(* IEC 61131-3 sources: SortJet_MasterSPS_Aufbau.fbsproj/09_Station/Stationen/_Basic/Basic_Schnittstelle_FB_V01_00_00.fb.st^, 6 files *)

(* ---- A_Changelog.act.st ---- *)
(* METADATA
{
	"v3Meta": {
		"objectGuid": "30bc6851-70b4-468b-8947-0ecaf15505c8"
	}
}
*)
{attribute 'excludefrombuild'}
ACTION A_Changelog
(* !!! VERSIONSÄNDERUNGEN WERDEN HIER DETAILLIERT DOKUMENTIERT !!!

- 2026-11-24 - V01_00_00: Tobias Brekerbohm
  - Erste Freigabe SortJet-Master
*)
END_ACTION

(* ---- A_Schnittstelle.act.st ---- *)
(* METADATA
{
	"v3Meta": {
		"objectGuid": "8ef5bc36-5f76-46e1-a5ac-606d922f719c"
	}
}
*)
ACTION A_Schnittstelle
//-------------------------------------------------------------------------------------------------
// AKTION SCHNITTSTELLE
//-------------------------------------------------------------------------------------------------

BasisStationsParameter.OutGlasTransport[cWAND_1].stStationsNummern          := BasisStationsParameter.stMKs.stStationsNummern;
BasisStationsParameter.OutGlasTransport[cWAND_1].wStationsTyp               := BasisStationsParameter.stMKs.eStationsTyp;
BasisStationsParameter.OutGlasTransport[cWAND_1].rLaengeStation             := BasisStationsParameter.stMKs.stFremdanlage.rLaengeStation;
BasisStationsParameter.OutGlasTransport[cWAND_1].bEinlaufsensor             REF= bEmpfaengerSensorEinlauf;
BasisStationsParameter.OutGlasTransport[cWAND_1].bAuslaufsensor             REF= bgFALSE;
BasisStationsParameter.OutGlasTransport[cWAND_1].bBereitZumAustransport     REF= blBereitZumAustransport;
BasisStationsParameter.OutGlasTransport[cWAND_1].bBereitZumEintransport     REF= blBereitZumEintransport;
BasisStationsParameter.OutGlasTransport[cWAND_1].rGeschwindigkeit           REF= rpGeschwindigkeit;
BasisStationsParameter.OutGlasTransport[cWAND_1].bFehler                    REF= BasisStationsParameter.bFehler;
BasisStationsParameter.OutGlasTransport[cWAND_1].bQuittScheibe              REF= bgFALSE;
BasisStationsParameter.OutGlasTransport[cWAND_1].bFreigabe                  REF= BasisStationsParameter.stFreigabe.bAlles;
BasisStationsParameter.OutGlasTransport[cWAND_1].bTransportAbgeschlossen    REF= bgFALSE;
BasisStationsParameter.OutGlasTransport[cWAND_1].bScheibeFaehrtUeberEinlauf REF= bgFALSE;
BasisStationsParameter.OutGlasTransport[cWAND_1].bScheibeFaehrtUeberAuslauf REF= bgFALSE;
BasisStationsParameter.OutGlasTransport[cWAND_1].bAutomatikBetriebAktiv     REF= blAutomatikBetriebAktiv;

//   - Status der Sortierung [Hardware- Ausgaenge]
//     => Automatik ativ
//     => Kein Fehler aktiv
out_bSenderBereit := blSenderBereit :=         BasisStationsParameter.bAutomatik
                     AND NOT BasisStationsParameter.bFehler
                     AND NOT BasisStationsParameter.InGlasTransportVorgaenger[cWAND_1].bFehler;

out_bSenderGlasBereit := blSenderGlasBereit (*OR bgVisu_Schnittstelle_GlasBereit[BasisStationsParameter.stMKs.stStationsNummern.NummerSPS]*);

// Eingangssignale können über den Drive oder IO's kommen
bEmpfaengerSensorEinlauf := bpEmpfaengerSensorEinlauf OR in_bEmpfaengerSensorEinlauf;

//-------------------------------------------------------------------------------------------------
// VISU
//-------------------------------------------------------------------------------------------------
bgVisu_Schnittstelle_GlasBereit[BasisStationsParameter.stMKs.stStationsNummern.NummerSPS]    := out_bSenderGlasBereit;
END_ACTION

(* ---- IGLineEvent.act.st ---- *)
(* METADATA
{
	"v3Meta": {
		"objectGuid": "eb410a9f-4f2d-4b91-9b42-1e80fc6ee1dd"
	}
}
*)
ACTION IGLineEvent
//-------------------------------------------------------------------------------------------------
// IG LINE EVENT
//-------------------------------------------------------------------------------------------------
bpISOLineEventAktiv := blUebergabeGlas;
(* Hinweis:
   - Ausgaenge setzen
*)
out_bLeuchteGlasbruch :=( blUebergabeGlas AND ((wpAuftragsTyp = 1) OR (wpAuftragsTyp = 4) OR ((wpAuftragsTyp = 5) AND gbFlashbit05sec))) ;
out_bLeuchteSpezial   :=( blUebergabeGlas AND ((wpAuftragsTyp = 2) OR ((wpAuftragsTyp = 3) AND gbFlashbit02sec )));

out_bAmpelEventAktiv := (blUebergabeGlas);

//-------------------------------------------------------------------------------------------------
// STEUERUNG:  ISO Line EVENT abhandeln
//-------------------------------------------------------------------------------------------------
IF ( bpStarteIGEvent
     AND NOT blUebergabeGlas )
THEN
  blUebergabeGlas := TRUE;
  bpStarteIGEvent := FALSE;
  steplUebergabeGlas := STEP_0_E;
END_IF

(* Hinweis:
   - wpAuftragsTyp:
   - case 0: //Kein Ereignis
   - case 1: //Scheibe von Isolinie abnehmen!
   - case 2: //Einschleusen von Sonderscheibe!
   - case 3: //Laufende!
   - case 4: //Alle Scheiben der Isoeinheit sind Bruch!
   - case 5: //Eine Scheibe der Einheit ist Bruch!
*)
IF ( blUebergabeGlas ) THEN
  CASE steplUebergabeGlas OF
    // GLASUEBERGABE ========================
    STEP_0_E:

      dwpWartezeit := 0;

      tlWarteZeiteAufnahme := TIME(); // Starten der Wartezeitenermittlung

      CASE wpAuftragsTyp OF
        0:
          steplUebergabeGlas:=STEP_1000_E;

        1,2,3,4,5:
          Horn.bpHornAktivieren := TRUE;
          Horn.wpStatusArt      := wpAuftragsTyp;
          Horn.tpHornZeit       := BasisStationsParameter.stMKs.stFremdanlage.tZeitHornAktiv;

          steplUebergabeGlas:=STEP_10_E;

        ELSE
          steplUebergabeGlas:=STEP_1000_E;
      END_CASE

    // GLASUEBERGABE ========================
    STEP_10_E:
      rtlTasterSpezial( CLK := in_bTasterSpezial );
      rtlTasterGlasbruch( CLK := in_bTasterGlasbruch );

      IF ((wpAuftragsTyp = 1) OR (wpAuftragsTyp = 4) OR (wpAuftragsTyp = 5))
         AND rtlTasterGlasbruch.CLK
      THEN
        steplUebergabeGlas:=STEP_100_E;
      END_IF

      IF ((wpAuftragsTyp = 2) OR (wpAuftragsTyp = 3))
         AND rtlTasterSpezial.Q
      THEN
        steplUebergabeGlas:=STEP_100_E;
      END_IF

    // GLASUEBERGABE ========================
    STEP_100_E:
      (* Hinweis:
         - Nachrichtabsetzen
      *)
      dwpWartezeit := TIME_TO_DWORD(TIME()- tlWarteZeiteAufnahme);
      wSps2MmiQuittISOLineNr   := BasisStationsParameter.stMKs.stStationsNummern.NummerIntern;
      dwSps2MmiWartezeit       := dwpWartezeit;
      MsgToMmi(auftragsnr_w    := SB0_SPS_SORTIERUNGQUITTUNGVONISOLINIE );

      steplUebergabeGlas:=STEP_1000_E;

    // GLASUEBERGABE ========================
    STEP_1000_E:
      steplUebergabeGlas:=STEP_0_E;
      blUebergabeGlas:=FALSE;
      dwpWartezeit := 0;

  // GLASUEBERGABE ========================
  END_CASE
END_IF

//-------------------------------------------------------------------------------------------------
// STEUERUNG: Abbruch eines ISO Line Events
//-------------------------------------------------------------------------------------------------
(* Hinweis:
   - Abbruch des ISO-Linie Event per MMI Nachricht [Cancel- Event]
   - Abbruch nach einem Stopp da das ISO-Linie Event nochmal geschickt wird
*)
IF ( bpResetISOLinieEvent ) THEN
  bpResetISOLinieEvent := FALSE;
  bpStarteIGEvent      := FALSE;
  blUebergabeGlas      := FALSE;
END_IF
END_ACTION

(* ---- M_GeschwindigkeitGlaetten.meth.st ---- *)
(* METADATA
{
	"v3Meta": {
		"objectGuid": "0474b6fd-4043-4228-8e53-82e27dbe01a7"
	}
}
*)
METHOD M_GeschwindigkeitGlaetten
VAR_INPUT
  rpMindestGeschwindigkeitsAenderung  : REAL; // MK stFremdanlage.rMindestGeschwindigkeitsAenderung
  tpMindestZeitZwischenGeschwAenderung : TIME; // MK stFremdanlage.tMindestZeitZwischenGeschwAenderung
END_VAR
VAR
  rlGeschwindigkeitSoll              : REAL; // Ungeglaettete Geschwindigkeit aus der Schnittstelle
  rlMindestGeschwindigkeitsAenderung : REAL;
END_VAR
//-------------------------------------------------------------------------------------------------
// GLAETTUNG: GESCHWINDIGKEIT ZUR SORTIERUNG
//-------------------------------------------------------------------------------------------------
(* Hinweis:
   - Aufruf in der abgeleiteten Schnittstelle, nachdem rpGeschwindigkeit berechnet wurde
   - Eine neue Geschwindigkeit wird nur uebernommen, wenn sie sich um mindestens
     rMindestGeschwindigkeitsAenderung geaendert hat und seit der letzten Uebernahme
     tMindestZeitZwischenGeschwAenderung vergangen ist
   - Stillstand (0) wird immer sofort ausgegeben, der erste Wert danach ebenfalls
*)
rlGeschwindigkeitSoll              := rpGeschwindigkeit;
rlMindestGeschwindigkeitsAenderung := MAX( rpMindestGeschwindigkeitsAenderung, 0.0 );

IF ( rlGeschwindigkeitSoll = 0.0 ) THEN
  rlGeschwindigkeitFreigegeben       := 0.0;
  blGeschwindigkeitInitialisiert     := FALSE;
  blGeschwindigkeitUpdateSperreAktiv := FALSE;

ELSIF NOT blGeschwindigkeitInitialisiert THEN
  rlGeschwindigkeitFreigegeben       := rlGeschwindigkeitSoll;
  blGeschwindigkeitInitialisiert     := TRUE;
  blGeschwindigkeitUpdateSperreAktiv := TRUE;

ELSIF NOT blGeschwindigkeitUpdateSperreAktiv
      AND ( ABS( rlGeschwindigkeitSoll - rlGeschwindigkeitFreigegeben ) >= rlMindestGeschwindigkeitsAenderung )
THEN
  rlGeschwindigkeitFreigegeben       := rlGeschwindigkeitSoll;
  blGeschwindigkeitUpdateSperreAktiv := TRUE;
END_IF

// Sperrzeit abgelaufen -> Aenderung ab dem naechsten Zyklus wieder freigeben
IF ( blGeschwindigkeitUpdateSperreAktiv AND tonlGeschwindigkeitUpdateSperre.Q ) THEN
  blGeschwindigkeitUpdateSperreAktiv := FALSE;
END_IF

tonlGeschwindigkeitUpdateSperre( IN := blGeschwindigkeitUpdateSperreAktiv,
                                 PT := tpMindestZeitZwischenGeschwAenderung );

rpGeschwindigkeit := rlGeschwindigkeitFreigegeben;
END_METHOD

(* ---- Meldungen.act.st ---- *)
(* METADATA
{
	"v3Meta": {
		"objectGuid": "44589f73-366e-43f4-b889-8e113549444f"
	}
}
*)
ACTION Meldungen
//-------------------------------------------------------------------------------------------------
// AKTION: MELDUNGEN
//-------------------------------------------------------------------------------------------------
// Meldungsnummer übergeben
wlWatchIONachrichtenNummer := BasisStationsParameter.stMKs.wMeldungsNummer;

WatchIoControl(T#30S ,wlWatchIONachrichtenNummer + 2  ,( blSenderBereit AND blSenderGlasBereit AND NOT blBereitZumEintransport));
END_ACTION

(* ---- Reset.act.st ---- *)
(* METADATA
{
	"v3Meta": {
		"objectGuid": "a6ec1752-3ec8-4f8b-95bc-dc8d5c4fd619"
	}
}
*)
ACTION Reset
//-------------------------------------------------------------------------------------------------
// AKTION: RESET
//-------------------------------------------------------------------------------------------------
AuftragsSpeicher( bpReset := TRUE );

blUebergabeGlas := FALSE;
wpAuftragsTyp := 0;
steplUebergabeGlas := STEP_0_E;

BasisStationsParameter.bCheckMitVorgaenger[cWAND_1] := FALSE;
BasisStationsParameter.bCheckMitNachfolger[cWAND_1] := FALSE;
BasisStationsParameter.bFehler                      := FALSE;
BasisStationsParameter.bAuftragAktiv                := FALSE;
BasisStationsParameter.bReset                       := FALSE;
END_ACTION
